(* ================================================================= *)
(*  FB_1020_EquipmentHandshake                                       *)
(*  通用设备通讯握手功能块 - 双通道状态机(与传输层无关)               *)
(*  版本: V2.0.0  日期: 2026-05-30                                    *)
(*  来源: SysLib/communication/                                      *)
(*  规范: LSP-905 V1.0.1, LSP-904 V1.2.0, LSP-903 V1.0.0            *)
(*                                                                    *)
(*  职责:                                                            *)
(*    - 上游送出握手: RequestOut -> Delay -> MoveBusy -> Complete     *)
(*    - 下游接收握手: RequestIn -> Delay -> MoveBusy -> Complete      *)
(*    - 双通道心跳监视 + 超时诊断                                     *)
(*    - 产品数据锁存透传(上升沿一次性锁存)                            *)
(*    - 接收侧产品数据输出                                            *)
(*                                                                    *)
(*  设计原则:                                                         *)
(*    - 纯协议逻辑, 不依赖任何具体传输层(Modbus/Profinet/OPC-UA等)     *)
(*    - 通过 VAR_IN_OUT io_stUpStream/io_stDownStream 与外部交换信号  *)
(*    - 信号映射由调用方(OB1)负责, 本FB只管时序和状态转换              *)
(*                                                                    *)
(*  V2.0.0 变更(Breaking Change):                                    *)
(*    - ST_ProductData: GlassID 30 INT -> 16 WORD                    *)
(*    - ST_HandshakeCh: 扁平字段 -> WriteProduct/ReadProduct 嵌入    *)
(*    - [B1] Disable段不再清除Write.Ready/DsReady/Reserved1-6        *)
(*    - [B2] 上游COMPLETE态增加Write.Complete回传                    *)
(*    - [B3] 产品数据改为MoveBusy上升沿一次性锁存                    *)
(*    - [D1] 新增q_stUpReceivedProduct/q_stDownReceivedProduct输出   *)
(*    - Disable段精简: 只清除FB管理的信号, 不触碰外部写入字段         *)
(*                                                                    *)
(*  协议来源: 各設備交握-5.20.xlsx 交握時序Sheet                      *)
(* ================================================================= *)

FUNCTION_BLOCK FB_1020_EquipmentHandshake

VAR_INPUT
    i_bEnable        : BOOL := FALSE;   // 使能 TRUE=执行握手逻辑
    i_bRequestOut    : BOOL := FALSE;   // 向上游发起要料请求
    i_bAllowDischarge: BOOL := FALSE;   // 允许向下游出料
    i_bReset         : BOOL := FALSE;   // 复位故障/强制回IDLE
    i_bTransportDone : BOOL := FALSE;   // 物理搬运完成信号(输送机构反馈)

    i_stProductData  : ST_ProductData;  // 待传递的产品跟踪数据

    i_dReqDelayMs    : DINT := 1000;    // 请求->搬运 延迟时间 ms
    i_dHbToggleMs    : DINT := 500;     // 心跳翻转周期 ms
    i_dHbTimeoutMs   : DINT := 3000;    // 心跳超时阈值 ms
    i_dCompleteMs    : DINT := 500;     // 完成脉冲宽度 ms
END_VAR

VAR_OUTPUT
    q_bUpReady       : BOOL := FALSE;   // 上游设备就绪综合信号
    q_bDownReady     : BOOL := FALSE;   // 下游设备就绪综合信号
    q_bUpComplete    : BOOL := FALSE;   // 上游送出完成脉冲
    q_bDownComplete  : BOOL := FALSE;   // 下游接收完成脉冲
    q_bAlarm         : BOOL := FALSE;   // 综合报警输出
    q_wStatusCode    : WORD := 16#0000; // 状态码 Hi=上游 Lo=下游

    q_iUpState       : INT := 0;        // 上游状态机当前状态
    q_iDownState     : INT := 0;        // 下游状态机当前状态

    q_stUpReceivedProduct   : ST_ProductData; // 从上游接收的产品数据
    q_stDownReceivedProduct : ST_ProductData; // 从下游接收的产品数据
END_VAR

VAR_IN_OUT
    io_stUpStream    : ST_HandshakeCh;  // 上游通道 Write=本机->上游 Read=上游->本机
    io_stDownStream  : ST_HandshakeCh;  // 下游通道 Write=本机->下游 Read=下游->本机
END_VAR

VAR
    // ===== 状态机 =====
    iUpState         : INT := 0;        // 上游状态 0=IDLE 1=REQ_OUT 2=MOVE_BUSY 3=COMPLETE 4=FAULT
    iDownState       : INT := 0;        // 下游状态 0=IDLE 1=REQ_IN 2=MOVE_BUSY 3=COMPLETE 4=FAULT

    // ===== 定时器 (两阶段调用: 先设IN/PT, 后集中调用) =====
    tReqOutDelay     : FB_TON;          // RequestOut -> MoveBusy 延迟
    tReqInDelay      : FB_TON;          // RequestIn -> 响应延迟
    tHbUpTimeout     : FB_TON;          // 上游心跳超时
    tHbDsTimeout     : FB_TON;          // 下游心跳超时
    tHbToggle        : FB_TON;          // 心跳翻转周期
    tCompletePulseUp : FB_TON;          // 上游完成脉冲宽度
    tCompletePulseDs : FB_TON;          // 下游完成脉冲宽度

    // ===== 边沿检测 (FB_R_TRIG参数名为IN, 非CLK) =====
    rTrigRequestOut  : FB_R_TRIG;       // i_bRequestOut上升沿
    rTrigRequestIn   : FB_R_TRIG;       // Read.RequestIn上升沿
    rTrigUpComplete  : FB_R_TRIG;       // Read.Complete上升沿
    rTrigDsComplete  : FB_R_TRIG;       // Read.DsComplete上升沿
    rTrigTransport   : FB_R_TRIG;       // i_bTransportDone上升沿
    rTrigMoveBusyUp  : FB_R_TRIG;       // Write.MoveBusy上升沿(产品数据锁存触发)
    rTrigMoveBusyDs  : FB_R_TRIG;       // Write.DsMoveBusy上升沿(产品数据锁存触发)

    // ===== 心跳监视辅助 =====
    bLastUpHbA       : BOOL := FALSE;   // 上周期上游Read.Heartbeat
    bLastUpHbB       : BOOL := FALSE;   // 上周期上游Read.RcvHeartbeat
    bLastDsHbA       : BOOL := FALSE;   // 上周期下游Read.RcvHeartbeat
    bLastDsHbB       : BOOL := FALSE;   // 上周期下游Read.Heartbeat
    bUpHbChanged     : BOOL := FALSE;   // 上游心跳翻转标志
    bDsHbChanged     : BOOL := FALSE;   // 下游心跳翻转标志

    // ===== 产品数据锁存标志 =====
    bUpDataLatched   : BOOL := FALSE;   // 上游产品数据已锁存
    bDsDataLatched   : BOOL := FALSE;   // 下游产品数据已锁存
END_VAR


(* ================================================================== *)
(*  Phase 1: 逻辑处理 - 设置定时器输入/状态机转换/边沿检测            *)
(* ================================================================== *)

(* ==================== 使能判断 ==================== *)
IF NOT i_bEnable THEN
    // [B1] 只清除FB管理的信号, 不触碰外部写入字段(Ready/DsReady/Reserved1-6)
    io_stUpStream.Write.Heartbeat    := FALSE;
    io_stUpStream.Write.RequestOut   := FALSE;
    io_stUpStream.Write.MoveBusy     := FALSE;
    io_stUpStream.Write.Complete     := FALSE;
    io_stUpStream.Write.RcvHeartbeat := FALSE;
    io_stUpStream.Write.RequestIn    := FALSE;
    io_stUpStream.Write.DsMoveBusy   := FALSE;
    io_stUpStream.Write.DsComplete   := FALSE;

    io_stDownStream.Write.Heartbeat    := FALSE;
    io_stDownStream.Write.RequestOut   := FALSE;
    io_stDownStream.Write.MoveBusy     := FALSE;
    io_stDownStream.Write.Complete     := FALSE;
    io_stDownStream.Write.RcvHeartbeat := FALSE;
    io_stDownStream.Write.RequestIn    := FALSE;
    io_stDownStream.Write.DsMoveBusy   := FALSE;
    io_stDownStream.Write.DsComplete   := FALSE;

    q_bUpReady := FALSE;
    q_bDownReady := FALSE;
    q_bUpComplete := FALSE;
    q_bDownComplete := FALSE;
    q_bAlarm := FALSE;
    q_wStatusCode := 16#0000;
    q_iUpState := 0;
    q_iDownState := 0;
    iUpState := 0;
    iDownState := 0;

    tReqOutDelay.IN := FALSE;
    tReqInDelay.IN := FALSE;
    tHbUpTimeout.IN := FALSE;
    tHbDsTimeout.IN := FALSE;
    tHbToggle.IN := FALSE;
    tCompletePulseUp.IN := FALSE;
    tCompletePulseDs.IN := FALSE;

ELSE

q_iUpState := iUpState;
q_iDownState := iDownState;


(* ==================== 心跳翻转生成 ==================== *)
tHbToggle.IN := NOT tHbToggle.Q;
tHbToggle.PT := i_dHbToggleMs;

io_stUpStream.Write.Heartbeat := tHbToggle.Q;
io_stDownStream.Write.RcvHeartbeat := tHbToggle.Q;


(* ==================== 心跳超时监视 ==================== *)

bUpHbChanged := (io_stUpStream.Read.Heartbeat <> bLastUpHbA)
             OR (io_stUpStream.Read.RcvHeartbeat <> bLastUpHbB);
bLastUpHbA := io_stUpStream.Read.Heartbeat;
bLastUpHbB := io_stUpStream.Read.RcvHeartbeat;

IF bUpHbChanged THEN
    tHbUpTimeout.IN := FALSE;
    io_stUpStream.HbTimeout := FALSE;
ELSE
    tHbUpTimeout.IN := TRUE;
END_IF;
tHbUpTimeout.PT := i_dHbTimeoutMs;

bDsHbChanged := (io_stDownStream.Read.RcvHeartbeat <> bLastDsHbA)
             OR (io_stDownStream.Read.Heartbeat <> bLastDsHbB);
bLastDsHbA := io_stDownStream.Read.RcvHeartbeat;
bLastDsHbB := io_stDownStream.Read.Heartbeat;

IF bDsHbChanged THEN
    tHbDsTimeout.IN := FALSE;
    io_stDownStream.HbTimeout := FALSE;
ELSE
    tHbDsTimeout.IN := TRUE;
END_IF;
tHbDsTimeout.PT := i_dHbTimeoutMs;

IF tHbUpTimeout.Q THEN
    io_stUpStream.HbTimeout := TRUE;
END_IF;
IF tHbDsTimeout.Q THEN
    io_stDownStream.HbTimeout := TRUE;
END_IF;


(* ==================== 就绪综合信号 ==================== *)
q_bUpReady := io_stUpStream.Read.Ready
              AND (NOT io_stUpStream.CommFault)
              AND (NOT io_stUpStream.HbTimeout);

q_bDownReady := io_stDownStream.Read.DsReady
               AND (NOT io_stDownStream.CommFault)
               AND (NOT io_stDownStream.HbTimeout);


(* ==================== 边沿检测 ==================== *)
rTrigRequestOut(IN := i_bRequestOut, Q => rTrigRequestOut.Q);
rTrigRequestIn(IN := io_stDownStream.Read.RequestIn, Q => rTrigRequestIn.Q);
rTrigUpComplete(IN := io_stUpStream.Read.Complete, Q => rTrigUpComplete.Q);
rTrigDsComplete(IN := io_stDownStream.Read.DsComplete, Q => rTrigDsComplete.Q);
rTrigTransport(IN := i_bTransportDone, Q => rTrigTransport.Q);
rTrigMoveBusyUp(IN := io_stUpStream.Write.MoveBusy, Q => rTrigMoveBusyUp.Q);
rTrigMoveBusyDs(IN := io_stDownStream.Write.DsMoveBusy, Q => rTrigMoveBusyDs.Q);


(* ==================== 上游状态机 ==================== *)
(* 协议时序: IDLE --[RequestOut+Ready]--> REQ_OUT --[1s]--> MOVE_BUSY
   --[对方Complete]--> COMPLETE --> IDLE
   任何态--[HbTimeout]--> FAULT *)

CASE iUpState OF
    0:
        (* IDLE: 空闲等待 *)
        io_stUpStream.Write.RequestOut := FALSE;
        io_stUpStream.Write.MoveBusy := FALSE;
        io_stUpStream.Write.Complete := FALSE;
        tReqOutDelay.IN := FALSE;
        tCompletePulseUp.IN := FALSE;
        bUpDataLatched := FALSE;

        IF rTrigRequestOut.Q AND q_bUpReady THEN
            iUpState := 1;
        END_IF;

        IF io_stUpStream.HbTimeout THEN
            iUpState := 4;
            io_stUpStream.CommFault := TRUE;
        END_IF;

    1:
        (* REQ_OUT: 已发出送料请求, 等待延迟 *)
        io_stUpStream.Write.RequestOut := TRUE;
        tReqOutDelay.IN := TRUE;
        tReqOutDelay.PT := i_dReqDelayMs;

        IF tReqOutDelay.Q THEN
            iUpState := 2;
            tReqOutDelay.IN := FALSE;
        END_IF;

        IF i_bReset OR io_stUpStream.HbTimeout THEN
            iUpState := 0;
            io_stUpStream.Write.RequestOut := FALSE;
            tReqOutDelay.IN := FALSE;
            IF io_stUpStream.HbTimeout THEN
                io_stUpStream.CommFault := TRUE;
            END_IF;
        END_IF;

    2:
        (* MOVE_BUSY_UP: 搬运中, 上升沿锁存产品数据 *)
        io_stUpStream.Write.MoveBusy := TRUE;
        io_stUpStream.Write.RequestOut := FALSE;

        (* [B3] MoveBusy上升沿一次性锁存产品数据 *)
        IF rTrigMoveBusyUp.Q AND (NOT bUpDataLatched) THEN
            io_stUpStream.WriteProduct := i_stProductData;
            bUpDataLatched := TRUE;
        END_IF;

        (* [D1] 上游Complete时锁存接收到的产品数据 *)
        IF rTrigUpComplete.Q THEN
            q_stUpReceivedProduct := io_stUpStream.ReadProduct;
            iUpState := 3;
        END_IF;

        IF i_bReset OR io_stUpStream.HbTimeout THEN
            iUpState := 0;
            io_stUpStream.Write.MoveBusy := FALSE;
            IF io_stUpStream.HbTimeout THEN
                io_stUpStream.CommFault := TRUE;
            END_IF;
        END_IF;

    3:
        (* COMPLETE_UP: [B2] 回传Complete + 完成脉冲后回IDLE *)
        io_stUpStream.Write.MoveBusy := FALSE;
        io_stUpStream.Write.Complete := TRUE;
        q_bUpComplete := TRUE;
        tCompletePulseUp.IN := TRUE;
        tCompletePulseUp.PT := i_dCompleteMs;

        IF tCompletePulseUp.Q THEN
            q_bUpComplete := FALSE;
            io_stUpStream.Write.Complete := FALSE;
            tCompletePulseUp.IN := FALSE;
            iUpState := 0;
        END_IF;

    4:
        (* FAULT_UP: 故障冻结, 等待复位或恢复 *)
        io_stUpStream.CommFault := TRUE;

        IF i_bReset OR (NOT io_stUpStream.HbTimeout) THEN
            io_stUpStream.CommFault := FALSE;
            io_stUpStream.Write.RequestOut := FALSE;
            io_stUpStream.Write.MoveBusy := FALSE;
            io_stUpStream.Write.Complete := FALSE;
            iUpState := 0;
        END_IF;

ELSE
    iUpState := 0;
END_CASE;


(* ==================== 下游状态机 ==================== *)
(* 协议时序: IDLE --[RequestIn+AllowDischarge+DownReady]--> REQ_IN --[1s]--> MOVE_BUSY
   --[TransportDone]--> COMPLETE --> IDLE
   任何态--[HbTimeout]--> FAULT *)

CASE iDownState OF
    0:
        (* IDLE: 空闲等待 *)
        io_stDownStream.Write.RequestIn := FALSE;
        io_stDownStream.Write.DsMoveBusy := FALSE;
        io_stDownStream.Write.DsComplete := FALSE;
        tReqInDelay.IN := FALSE;
        tCompletePulseDs.IN := FALSE;
        bDsDataLatched := FALSE;

        IF rTrigRequestIn.Q AND i_bAllowDischarge AND q_bDownReady THEN
            iDownState := 1;
        END_IF;

        IF io_stDownStream.HbTimeout THEN
            iDownState := 4;
            io_stDownStream.CommFault := TRUE;
        END_IF;

    1:
        (* REQ_IN: 收到请求, 等待响应延迟 *)
        tReqInDelay.IN := TRUE;
        tReqInDelay.PT := i_dReqDelayMs;

        IF tReqInDelay.Q THEN
            iDownState := 2;
            tReqInDelay.IN := FALSE;
        END_IF;

        IF i_bReset OR io_stDownStream.HbTimeout
           OR (NOT io_stDownStream.Read.RequestIn) THEN
            iDownState := 0;
            tReqInDelay.IN := FALSE;
            IF io_stDownStream.HbTimeout THEN
                io_stDownStream.CommFault := TRUE;
            END_IF;
        END_IF;

    2:
        (* MOVE_BUSY_DS: 搬运中, 上升沿锁存产品数据, 等待物理传输完成 *)
        io_stDownStream.Write.DsMoveBusy := TRUE;

        (* [B3] DsMoveBusy上升沿一次性锁存产品数据 *)
        IF rTrigMoveBusyDs.Q AND (NOT bDsDataLatched) THEN
            io_stDownStream.WriteProduct := i_stProductData;
            bDsDataLatched := TRUE;
        END_IF;

        IF rTrigTransport.Q OR rTrigDsComplete.Q THEN
            (* [D1] 锁存下游接收到的产品数据 *)
            q_stDownReceivedProduct := io_stDownStream.ReadProduct;
            iDownState := 3;
        END_IF;

        IF i_bReset OR io_stDownStream.HbTimeout THEN
            iDownState := 0;
            io_stDownStream.Write.DsMoveBusy := FALSE;
            IF io_stDownStream.HbTimeout THEN
                io_stDownStream.CommFault := TRUE;
            END_IF;
        END_IF;

    3:
        (* COMPLETE_DS: 完成脉冲后回IDLE *)
        io_stDownStream.Write.DsMoveBusy := FALSE;
        io_stDownStream.Write.DsComplete := TRUE;
        q_bDownComplete := TRUE;
        tCompletePulseDs.IN := TRUE;
        tCompletePulseDs.PT := i_dCompleteMs;

        IF tCompletePulseDs.Q THEN
            q_bDownComplete := FALSE;
            io_stDownStream.Write.DsComplete := FALSE;
            tCompletePulseDs.IN := FALSE;
            iDownState := 0;
        END_IF;

    4:
        (* FAULT_DS: 故障冻结 *)
        io_stDownStream.CommFault := TRUE;

        IF i_bReset OR (NOT io_stDownStream.HbTimeout) THEN
            io_stDownStream.CommFault := FALSE;
            io_stDownStream.Write.RequestIn := FALSE;
            io_stDownStream.Write.DsMoveBusy := FALSE;
            io_stDownStream.Write.DsComplete := FALSE;
            iDownState := 0;
        END_IF;

ELSE
    iDownState := 0;
END_CASE;


(* ==================== 综合报警 ==================== *)
q_bAlarm := io_stUpStream.CommFault OR io_stDownStream.CommFault
           OR io_stUpStream.HbTimeout OR io_stDownStream.HbTimeout;

(* ==================== 状态码 ==================== *)
q_wStatusCode := SHL(INT_TO_WORD(iUpState), 8) OR INT_TO_WORD(iDownState);


END_IF;

(* ================================================================== *)
(*  Phase 2: 定时器集中调用 - 将IN/PT传入, Q/ET输出回自身成员        *)
(*  必须每个扫描周期都调用, 否则定时器内部状态不更新                   *)
(* ================================================================== *)

tHbToggle(IN := tHbToggle.IN, PT := tHbToggle.PT,
          Q => tHbToggle.Q, ET => tHbToggle.ET);

tHbUpTimeout(IN := tHbUpTimeout.IN, PT := tHbUpTimeout.PT,
             Q => tHbUpTimeout.Q, ET => tHbUpTimeout.ET);

tHbDsTimeout(IN := tHbDsTimeout.IN, PT := tHbDsTimeout.PT,
             Q => tHbDsTimeout.Q, ET => tHbDsTimeout.ET);

tReqOutDelay(IN := tReqOutDelay.IN, PT := tReqOutDelay.PT,
             Q => tReqOutDelay.Q, ET => tReqOutDelay.ET);

tReqInDelay(IN := tReqInDelay.IN, PT := tReqInDelay.PT,
            Q => tReqInDelay.Q, ET => tReqInDelay.ET);

tCompletePulseUp(IN := tCompletePulseUp.IN, PT := tCompletePulseUp.PT,
                 Q => tCompletePulseUp.Q, ET => tCompletePulseUp.ET);

tCompletePulseDs(IN := tCompletePulseDs.IN, PT := tCompletePulseDs.PT,
                 Q => tCompletePulseDs.Q, ET => tCompletePulseDs.ET);

END_FUNCTION_BLOCK
